FUNCTION_BLOCK FB_CC_TempSensor EXTENDS FB_TempSensor_FFO
VAR
    rtVetoReset: R_TRIG;
END_VAR

// Reset the FFO for transitions to bVeto
// bAutoreset is False, but we still want to clear the fault on veto
rtVetoReset(CLK:=bVeto);
FFO.i_xReset := rtVetoReset.Q;

SUPER^(bAutoReset:=FALSE, io_fbFFHWO:=io_fbFFHWO);

END_FUNCTION_BLOCK

(* stored: Version 1.1.0.1
   POU FB_CC_TempSensor: Id {62e52992-2558-4a9c-b1dd-b3b9616cbbcf}, SpecialFunc None *)
